// TwinCAT 3 PLC project StateMachineControl
// ProgramVersion: 3.1.4026.22
// libraries:
//   Tc2_Standard, * (Beckhoff Automation GmbH)
//   Tc2_System, * (Beckhoff Automation GmbH)
// project tree:
//   DUTs/ E_DriveState.TcDUT, E_ModeState.TcDUT, ST_ModeOutputs.TcDUT, ST_ModeManagerActions.TcDUT
//   GVLs/ GVL_MODE.TcGVL
//   / PlcTask.TcTTO
//   POUs/ FB_StateMachineControl.TcPOU, FB_HeartbeatWatchdog.TcPOU, FB_ModeManagerCore.TcPOU, F_DeriveModeOutputs.TcPOU, MAIN.TcPOU, F_DecodeDriveState.TcPOU
// real-time tasks:
//   TASK VirtualMotorTask: cycle T#125us, priority 1, ADS port 351
//   TASK StateTask: cycle T#10ms, priority 2, ADS port 355
// variable links:
//   ExperimentSequencer/ExperimentSequencer Instance <-> StateMachineControl/StateMachineControl Instance
//     VirtualMotorTask Inputs/GVL_SEQ.experimentActive <-> PlcTask Outputs/MAIN.experimentActiveOut
//     VirtualMotorTask Inputs/GVL_SEQ.resetReq <-> PlcTask Outputs/MAIN.resetOut
//     VirtualMotorTask Outputs/GVL_SEQ.playbackDone <-> PlcTask Inputs/MAIN.seqPlaybackDone
//   ExperimentSequencer/ExperimentSequencer Instance <-> ControllerCore/ControllerCore_Obj1 (Module1)
//     VirtualMotorTask Outputs/GVL_SEQ.ffValue <-> Inputs/ffValue
//     VirtualMotorTask Outputs/GVL_SEQ.refValue <-> Inputs/refValue
//   ExperimentSequencer/ExperimentSequencer Instance <-> DriverAdapter/DriverAdapter_Obj1 (Module1)
//     VirtualMotorTask Outputs/GVL_SEQ.distValue <-> Inputs/distValue
//     VirtualMotorTask Outputs/GVL_SEQ.playbackDone <-> Inputs/playbackDone
//   ExperimentSequencer/ExperimentSequencer Instance <-> ExperimentLogger/ExperimentLogger_Obj1 (Module1)
//     VirtualMotorTask Outputs/GVL_SEQ.distValue <-> Inputs/record/distValue
//     VirtualMotorTask Outputs/GVL_SEQ.ffValue <-> Inputs/record/ffValue
//     VirtualMotorTask Outputs/GVL_SEQ.playbackDone <-> Inputs/control/playbackDone
//     VirtualMotorTask Outputs/GVL_SEQ.refValue <-> Inputs/record/refValue
//   StateMachineControl/StateMachineControl Instance <-> ControllerCore/ControllerCore_Obj1 (Module1)
//     PlcTask Outputs/MAIN.resetOut <-> Inputs/resetReq
//   StateMachineControl/StateMachineControl Instance <-> DriverAdapter/DriverAdapter_Obj1 (Module1)
//     PlcTask Inputs/MAIN.loadStatWord <-> Outputs/loadStatusWordOut
//     PlcTask Inputs/MAIN.motorStatWord <-> Outputs/motorStatusWordOut
//     PlcTask Outputs/MAIN.enableCurrentOut <-> Inputs/enableCurrentOutput
//     PlcTask Outputs/MAIN.loadCtrlWord <-> Inputs/loadControlWordIn
//     PlcTask Outputs/MAIN.motorCtrlWord <-> Inputs/motorControlWordIn
//     PlcTask Outputs/MAIN.resetOut <-> Inputs/resetReq
//   StateMachineControl/StateMachineControl Instance <-> ExperimentLogger/ExperimentLogger_Obj1 (Module1)
//     PlcTask Inputs/MAIN.loggerErrorCodeIn <-> Outputs/status/errorCode
//     PlcTask Inputs/MAIN.loggerFileReleasedIn <-> Outputs/status/fileReleased
//     PlcTask Inputs/MAIN.loggerReadyIn <-> Outputs/status/loggerReady
//     PlcTask Outputs/MAIN.experimentActiveOut <-> Inputs/control/loggingReq
//     PlcTask Outputs/MAIN.preArmOut <-> Inputs/control/preArmReq
//     PlcTask Outputs/MAIN.resetOut <-> Inputs/control/resetReq
//   ControllerCore/ControllerCore_Obj1 (Module1) <-> DriverAdapter/DriverAdapter_Obj1 (Module1)
//     Inputs/positionAct <-> Outputs/load/positionRel
//     Outputs/controlInput <-> Inputs/controlInput
//   ControllerCore/ControllerCore_Obj1 (Module1) <-> ExperimentLogger/ExperimentLogger_Obj1 (Module1)
//     Outputs/controlInput <-> Inputs/record/controlInput
//     Outputs/error <-> Inputs/record/error
//   DriverAdapter/DriverAdapter_Obj1 (Module1) <-> ExperimentLogger/ExperimentLogger_Obj1 (Module1)
//     Outputs/currentCmd <-> Inputs/record/currentCmd
//     Outputs/load/positionRel <-> Inputs/record/load/position
//     Outputs/load/velocityAct <-> Inputs/record/load/velocity
//     Outputs/motor/currentAct <-> Inputs/record/motor/currentAct
//     Outputs/motor/positionRel <-> Inputs/record/motor/position
//     Outputs/motor/velocityAct <-> Inputs/record/motor/velocity
//   DriverAdapter/DriverAdapter_Obj1 (Module1) <-> RealMotorPdo/RealMotorPdo Instance
//     Inputs/loadRaw/positionActualValue <-> Outputs/load/positionActualValue
//     Inputs/loadRaw/statusWord <-> Outputs/load/statusWord
//     Inputs/loadRaw/torqueActualValue <-> Outputs/load/torqueActualValue
//     Inputs/loadRaw/velocityActualValue <-> Outputs/load/velocityActualValue
//     Inputs/motorRaw/positionActualValue <-> Outputs/motor/positionActualValue
//     Inputs/motorRaw/statusWord <-> Outputs/motor/statusWord
//     Inputs/motorRaw/torqueActualValue <-> Outputs/motor/torqueActualValue
//     Inputs/motorRaw/velocityActualValue <-> Outputs/motor/velocityActualValue
//     Outputs/loadControlWordOut <-> Inputs/load/controlWord
//     Outputs/motorControlWordOut <-> Inputs/motor/controlWord
//     Outputs/targetTorque <-> Inputs/motor/targetTorque

CONFIGURATION StateMachineControl
    RESOURCE PLC ON TwinCAT3
        TASK PlcTask(INTERVAL := T#10ms, PRIORITY := 2);
        PROGRAM MAIN WITH PlcTask : MAIN;
    END_RESOURCE
END_CONFIGURATION

// ---- DUTs/E_DriveState.TcDUT
{attribute 'qualified_only'}
{attribute 'strict'}
{attribute 'to_string'}
TYPE E_DriveState :
(
    UNKNOWN := 0,

    // CiA402 "Switch on disabled"
    SWITCH_ON_DISABLED := 10,

    // CiA402 "Ready to switch on"
    READY_TO_SWITCH_ON := 20,

    // CiA402 "Switched on"
    SWITCHED_ON := 30,

    // CiA402 "Operation enabled"
    OPERATION_ENABLED := 40,

    // CiA402 "Fault"
    FAULT := 90
);
END_TYPE

// ---- DUTs/E_ModeState.TcDUT
{attribute 'qualified_only'}
{attribute 'strict'}
{attribute 'to_string'}
TYPE E_ModeState :
(
    IDLE := 0,              // Servo OFF / initial
    RESETTING := 10,        // Reset pulse active — no experiment transitions allowed
    SERVO_READY := 20,      // Servo ON + drive OPERATION_ENABLED, awaiting experiment
    RUNNING := 30,          // Experiment active
    DONE := 40              // Playback complete, awaiting rearm
);
END_TYPE

// ---- DUTs/ST_ModeOutputs.TcDUT
TYPE ST_ModeOutputs :
STRUCT
    experimentActiveOut : BOOL;
    preArmOut : BOOL;
    resetOut : BOOL;
    enableCurrentOut : BOOL;
END_STRUCT
END_TYPE

// ---- DUTs/ST_ModeManagerActions.TcDUT
TYPE ST_ModeManagerActions :
STRUCT
    consumeResetReq : BOOL;
    clearModeFlags : BOOL;
    incrementResetAckCounter : BOOL;
    incrementWatchdogTripCounter : BOOL;
END_STRUCT
END_TYPE

// ---- GVLs/GVL_MODE.TcGVL
{attribute 'qualified_only'}
VAR_GLOBAL CONSTANT
    MODEF_SERVO_ENABLE : UINT := 16#0001;          (* bit0 *)
    MODEF_EXPERIMENT_START_REQ : UINT := 16#0002;  (* bit1 *)
    HEARTBEAT_TIMEOUT_TICKS : UDINT := 50;         (* 10 ms task * 50 = 500 ms *)

END_VAR

VAR_GLOBAL
    {attribute 'linkalways'}
    modeFlags : UINT := 0;
    resetReq : BOOL := FALSE;
    resetAckCounter : UDINT := 0;
    hostHeartbeatCounter : UDINT := 0;
    watchdogTripCounter : UDINT := 0;
    experimentActive : BOOL := FALSE;
    loggerFileReleased : BOOL := FALSE;
    loggerErrorCode : UDINT := 0;
    modeState : E_ModeState := E_ModeState.IDLE;
END_VAR

// ---- POUs/MAIN.TcPOU
PROGRAM MAIN
VAR
    motorCtrlWord AT%Q* : UINT; // Motor ControlWord output
    loadCtrlWord AT%Q* : UINT; // Load ControlWord output
    motorStatWord AT%I* : UINT; // Motor StatusWord input
    loadStatWord AT%I* : UINT; // Load StatusWord input
    seqPlaybackDone AT%I* : BOOL; // Sequencer playback done (latched)
    experimentActiveOut AT%Q* : BOOL; // ModeManager experiment active output
    preArmOut AT%Q* : BOOL; // ModeManager logger pre-arm output
    resetOut AT%Q* : BOOL; // One-shot reset pulse output
    enableCurrentOut AT%Q* : BOOL; // Current enable gate output

    // FSM state
    modeState : E_ModeState := E_ModeState.IDLE;
    modeOutputs : ST_ModeOutputs;

    // Decoded request flags (from GVL_MODE.modeFlags)
    servoEnableReq : BOOL := FALSE;
    experimentStartReq : BOOL := FALSE;
    fbModeManagerCore : FB_ModeManagerCore;

    // Drive state
    driveReady : BOOL := FALSE;
    motorDriveReady : BOOL := FALSE;
    loadDriveReady : BOOL := FALSE;
    enableEffective : BOOL := FALSE;

    fbMotorStateMachine : FB_StateMachineControl;
    fbLoadStateMachine : FB_StateMachineControl;
    loggerReadyIn AT%I* : BOOL; // ExperimentLogger file FSM ACTIVE
    loggerFileReleasedIn AT%I* : BOOL; // ExperimentLogger close completed
    loggerErrorCodeIn AT%I* : UDINT; // ExperimentLogger session error
END_VAR

(* ===== 1. Decode input flags ===== *)
servoEnableReq := (GVL_MODE.modeFlags AND GVL_MODE.MODEF_SERVO_ENABLE) <> 0;
experimentStartReq := (GVL_MODE.modeFlags AND GVL_MODE.MODEF_EXPERIMENT_START_REQ) <> 0;

(* ===== 2. Request/watchdog/FSM core ===== *)
fbModeManagerCore(
    servoEnableRequest := servoEnableReq,
    experimentStartRequest := experimentStartReq,
    anyModeRequest := (GVL_MODE.modeFlags <> 0),
    resetRequest := GVL_MODE.resetReq,
    experimentActivePreviousScan := GVL_MODE.experimentActive,
    hostHeartbeatCounter := GVL_MODE.hostHeartbeatCounter,
    heartbeatTimeoutTicks := GVL_MODE.HEARTBEAT_TIMEOUT_TICKS,
    driveReadyPreviousScan := driveReady,
    loggerReady := loggerReadyIn,
    seqPlaybackDone := seqPlaybackDone
);

IF fbModeManagerCore.actions.consumeResetReq THEN
    GVL_MODE.resetReq := FALSE;
END_IF
IF fbModeManagerCore.actions.clearModeFlags THEN
    GVL_MODE.modeFlags := 0;
END_IF
IF fbModeManagerCore.actions.incrementResetAckCounter THEN
    GVL_MODE.resetAckCounter := GVL_MODE.resetAckCounter + 1;
END_IF
IF fbModeManagerCore.actions.incrementWatchdogTripCounter THEN
    GVL_MODE.watchdogTripCounter := GVL_MODE.watchdogTripCounter + 1;
END_IF

modeState := fbModeManagerCore.modeState;
enableEffective := fbModeManagerCore.driveEnable;

(* ===== 3. Drive state update ===== *)
fbMotorStateMachine(
    statusWord := motorStatWord,
    enable := enableEffective
);
fbLoadStateMachine(
    statusWord := loadStatWord,
    enable := enableEffective
);

motorCtrlWord := fbMotorStateMachine.controlWord;
loadCtrlWord := fbLoadStateMachine.controlWord;
motorDriveReady := (fbMotorStateMachine.driveState = E_DriveState.OPERATION_ENABLED);
loadDriveReady := (fbLoadStateMachine.driveState = E_DriveState.OPERATION_ENABLED);
driveReady := motorDriveReady AND loadDriveReady;

(* ===== 4. State-dependent outputs ===== *)
modeOutputs := F_DeriveModeOutputs(modeState := modeState);
experimentActiveOut := modeOutputs.experimentActiveOut;
preArmOut := modeOutputs.preArmOut;
resetOut := modeOutputs.resetOut;
enableCurrentOut := modeOutputs.enableCurrentOut;

GVL_MODE.experimentActive := experimentActiveOut;
IF modeState = E_ModeState.SERVO_READY THEN
    GVL_MODE.loggerFileReleased := FALSE;
    GVL_MODE.loggerErrorCode := 0;
ELSE
    GVL_MODE.loggerFileReleased := loggerFileReleasedIn;
    GVL_MODE.loggerErrorCode := loggerErrorCodeIn;
END_IF;
GVL_MODE.modeState := modeState;

END_PROGRAM

// ---- POUs/FB_ModeManagerCore.TcPOU
FUNCTION_BLOCK FB_ModeManagerCore
VAR_INPUT
    servoEnableRequest : BOOL;
    experimentStartRequest : BOOL;
    anyModeRequest : BOOL;
    resetRequest : BOOL;
    experimentActivePreviousScan : BOOL;
    hostHeartbeatCounter : UDINT;
    heartbeatTimeoutTicks : UDINT;
    driveReadyPreviousScan : BOOL;
    loggerReady : BOOL;
    seqPlaybackDone : BOOL;
END_VAR
VAR_OUTPUT
    modeState : E_ModeState := E_ModeState.IDLE;
    driveEnable : BOOL := FALSE;
    watchdogArmed : BOOL := FALSE;
    watchdogTimeout : BOOL := FALSE;
    actions : ST_ModeManagerActions;
END_VAR
VAR
    servoEnableRequestPrev : BOOL := FALSE;
    experimentStartRequestPrev : BOOL := FALSE;
    servoEnableEdge : BOOL := FALSE;
    experimentStartEdge : BOOL := FALSE;
    servoEnableLatched : BOOL := FALSE;
    experimentStartLatched : BOOL := FALSE;
    resetRequestPrev : BOOL := FALSE;
    resetEdge : BOOL := FALSE;
    resetHoldTicksRemaining : UDINT := 0;
    fbHeartbeatWatchdog : FB_HeartbeatWatchdog;
END_VAR
VAR CONSTANT
    RESET_PULSE_HOLD_TICKS : UDINT := 1;
END_VAR

actions.consumeResetReq := FALSE;
actions.clearModeFlags := FALSE;
actions.incrementResetAckCounter := FALSE;
actions.incrementWatchdogTripCounter := FALSE;

servoEnableEdge := servoEnableRequest AND NOT servoEnableRequestPrev;
experimentStartEdge := experimentStartRequest AND NOT experimentStartRequestPrev;
servoEnableRequestPrev := servoEnableRequest;
experimentStartRequestPrev := experimentStartRequest;

IF servoEnableEdge THEN
    servoEnableLatched := TRUE;
END_IF
IF experimentStartEdge THEN
    experimentStartLatched := TRUE;
END_IF
(* A missing servo request is the explicit abort contract.  Clear both
   latches so a start captured during RESETTING cannot run after rearm. *)
IF NOT servoEnableRequest THEN
    servoEnableLatched := FALSE;
    experimentStartLatched := FALSE;
END_IF

resetEdge := resetRequest AND NOT resetRequestPrev;
IF resetEdge THEN
    actions.consumeResetReq := TRUE;
END_IF
resetRequestPrev := resetRequest;

watchdogArmed := anyModeRequest OR experimentActivePreviousScan OR servoEnableLatched;
fbHeartbeatWatchdog(
    enable := watchdogArmed,
    heartbeatCounter := hostHeartbeatCounter,
    timeoutTicks := heartbeatTimeoutTicks
);
watchdogTimeout := fbHeartbeatWatchdog.timeout;

IF watchdogTimeout THEN
    modeState := E_ModeState.IDLE;
    actions.clearModeFlags := TRUE;
    servoEnableLatched := FALSE;
    experimentStartLatched := FALSE;
    IF fbHeartbeatWatchdog.tripEdge THEN
        actions.incrementWatchdogTripCounter := TRUE;
    END_IF

ELSIF resetEdge THEN
    modeState := E_ModeState.RESETTING;
    resetHoldTicksRemaining := RESET_PULSE_HOLD_TICKS;
    actions.clearModeFlags := TRUE;
    actions.incrementResetAckCounter := TRUE;
    servoEnableLatched := FALSE;
    experimentStartLatched := FALSE;

ELSE
    CASE modeState OF
        E_ModeState.IDLE:
            IF servoEnableLatched THEN
                modeState := E_ModeState.SERVO_READY;
            END_IF

        E_ModeState.RESETTING:
            IF resetHoldTicksRemaining > 0 THEN
                resetHoldTicksRemaining := resetHoldTicksRemaining - 1;
            ELSE
                modeState := E_ModeState.IDLE;
            END_IF

        E_ModeState.SERVO_READY:
            IF NOT servoEnableLatched THEN
                modeState := E_ModeState.IDLE;
                experimentStartLatched := FALSE;
            ELSIF experimentStartLatched AND driveReadyPreviousScan AND loggerReady THEN
                modeState := E_ModeState.RUNNING;
                experimentStartLatched := FALSE;
            END_IF

        E_ModeState.RUNNING:
            IF NOT servoEnableLatched OR NOT driveReadyPreviousScan THEN
                modeState := E_ModeState.IDLE;
                experimentStartLatched := FALSE;
                servoEnableLatched := FALSE;
                actions.clearModeFlags := TRUE;
            ELSIF seqPlaybackDone THEN
                modeState := E_ModeState.DONE;
                servoEnableLatched := FALSE;
                experimentStartLatched := FALSE;
                actions.clearModeFlags := TRUE;
            END_IF

        E_ModeState.DONE:
            servoEnableLatched := FALSE;
            experimentStartLatched := FALSE;
    END_CASE
END_IF

driveEnable := servoEnableLatched
    AND (modeState = E_ModeState.SERVO_READY OR modeState = E_ModeState.RUNNING);

END_FUNCTION_BLOCK

// ---- POUs/FB_HeartbeatWatchdog.TcPOU
FUNCTION_BLOCK FB_HeartbeatWatchdog
VAR_INPUT
    enable : BOOL;
    heartbeatCounter : UDINT;
    timeoutTicks : UDINT;
END_VAR
VAR_OUTPUT
    timeout : BOOL := FALSE;
    tripEdge : BOOL := FALSE;
END_VAR
VAR
    counterPrev : UDINT := 0;
    silenceTicks : UDINT := 0;
    tripLatched : BOOL := FALSE;
    heartbeatChanged : BOOL := FALSE;
END_VAR

tripEdge := FALSE;
heartbeatChanged := (heartbeatCounter <> counterPrev);

IF NOT enable THEN
    counterPrev := heartbeatCounter;
    silenceTicks := 0;
    tripLatched := FALSE;
ELSIF heartbeatChanged THEN
    counterPrev := heartbeatCounter;
    silenceTicks := 0;
    tripLatched := FALSE;
ELSE
    IF silenceTicks < timeoutTicks THEN
        silenceTicks := silenceTicks + 1;
    END_IF
END_IF

timeout := enable AND (silenceTicks >= timeoutTicks);
IF timeout AND NOT tripLatched THEN
    tripEdge := TRUE;
    tripLatched := TRUE;
END_IF

END_FUNCTION_BLOCK

// ---- POUs/FB_StateMachineControl.TcPOU
FUNCTION_BLOCK FB_StateMachineControl
VAR_INPUT
    statusWord : UINT; // 0x6041
    enable      : BOOL := TRUE;
END_VAR
VAR_OUTPUT
    controlWord : UINT;      // 0x6040
    driveState   : E_DriveState;
END_VAR
VAR
    faultResetPulsed : BOOL := FALSE;
END_VAR
VAR CONSTANT
    // Common CiA402 control commands (0x6040)
    CW_DISABLE_VOLTAGE : UINT := 16#0000;
    CW_SHUTDOWN        : UINT := 16#0006;
    CW_SWITCH_ON       : UINT := 16#0007;
    CW_ENABLE_OP       : UINT := 16#000F;
    CW_FAULT_RESET     : UINT := 16#0080;
END_VAR

driveState := F_DecodeDriveState(statusWord);

// Disable requested: force safe output
IF NOT enable THEN
    controlWord := CW_DISABLE_VOLTAGE;
    faultResetPulsed := FALSE;
    RETURN;
END_IF

CASE driveState OF

    E_DriveState.FAULT:
        // Fault reset should be a pulse. One scan is usually enough.
        IF NOT faultResetPulsed THEN
            controlWord := CW_FAULT_RESET;
            faultResetPulsed := TRUE;
        ELSE
            controlWord := CW_DISABLE_VOLTAGE;
        END_IF

    E_DriveState.SWITCH_ON_DISABLED:
        controlWord := CW_SHUTDOWN;
        faultResetPulsed := FALSE;

    E_DriveState.READY_TO_SWITCH_ON:
        controlWord := CW_SWITCH_ON;
        faultResetPulsed := FALSE;

    E_DriveState.SWITCHED_ON:
        controlWord := CW_ENABLE_OP;
        faultResetPulsed := FALSE;

    E_DriveState.OPERATION_ENABLED:
        controlWord := CW_ENABLE_OP;
        faultResetPulsed := FALSE;

    ELSE
        // UNKNOWN: converge from below (safe)
        controlWord := CW_SHUTDOWN;
        faultResetPulsed := FALSE;
END_CASE

END_FUNCTION_BLOCK

// ---- POUs/F_DecodeDriveState.TcPOU
FUNCTION F_DecodeDriveState : E_DriveState
VAR_INPUT
    statusWord : UINT; // 0x6041
END_VAR
VAR
    masked : UINT;
END_VAR

masked := statusWord AND 16#006F;

IF (masked AND 16#0008) <> 0 THEN
    // bit3 = Fault
    F_DecodeDriveState := E_DriveState.FAULT;
ELSIF masked = 16#0060 THEN
    // Switch on disabled
    F_DecodeDriveState := E_DriveState.SWITCH_ON_DISABLED;
ELSIF masked = 16#0021 THEN
    // Ready to switch on
    F_DecodeDriveState := E_DriveState.READY_TO_SWITCH_ON;
ELSIF masked = 16#0023 THEN
    // Switched on
    F_DecodeDriveState := E_DriveState.SWITCHED_ON;
ELSIF masked = 16#0027 THEN
    // Operation enabled
    F_DecodeDriveState := E_DriveState.OPERATION_ENABLED;
ELSE
    F_DecodeDriveState := E_DriveState.UNKNOWN;
END_IF

END_FUNCTION

// ---- POUs/F_DeriveModeOutputs.TcPOU
FUNCTION F_DeriveModeOutputs : ST_ModeOutputs
VAR_INPUT
    modeState : E_ModeState;
END_VAR

(* Safe default for unknown or newly added states. *)
F_DeriveModeOutputs.experimentActiveOut := FALSE;
F_DeriveModeOutputs.preArmOut := FALSE;
F_DeriveModeOutputs.resetOut := FALSE;
F_DeriveModeOutputs.enableCurrentOut := FALSE;

CASE modeState OF
    E_ModeState.RESETTING:
        F_DeriveModeOutputs.resetOut := TRUE;

    E_ModeState.SERVO_READY:
        F_DeriveModeOutputs.preArmOut := TRUE;
        F_DeriveModeOutputs.enableCurrentOut := TRUE;

    E_ModeState.RUNNING:
        F_DeriveModeOutputs.experimentActiveOut := TRUE;
        F_DeriveModeOutputs.enableCurrentOut := TRUE;
END_CASE

END_FUNCTION
